PROGRAM MAIN
VAR

	fTotalCIP_Volume: REAL;
	fbWritePersistent: FB_WritePersistentData;
	bTesting		:	BOOL:=FALSE	;
	nI_1			: 	INT		;
	ftg_EStop_Fall	: 	F_TRIG	;
	rs_EStopFall	: 	RS	;
	bTestEstop		:	BOOL:=TRUE	;
	bTemp_Water_Overweight_check: BOOL;
	fbUPS: FB_S_UPS_CX51x0;

END_VAR

prg_RealClock();
prg_Piston();
prg_Safety();
prg_MessageManager();
prg_Messages();
prg_Call_OpMode();
prg_User();
act_ResetPumps();
(*
prg_TriBlender(
		fb_TriBlenderPump:= g_Pump.fbPump[E_Pump_List.TB0001],
		stTriblender:=stTriblender,
		arrComponents:=arrProductionComponents);
*)		
//act_SetAnalogSens_Test();//To be deleted, for testing purposes
act_Call_Sensors_Analog();//To be deleted, for testing purposes
act_Call_Sensors_Analog_1();//To be deleted, for testing purposes
act_Call_ScaleFactor();//To be deleted, for testing purposes
act_Call_ProcessCntrl();

act_Call_Pumps();
act_Sensors();
act_HeatExchenger();
//CIP <-> Siemens exchange
g_Anybus.fbSim(arToCip:=g_Anybus.arSimRaw, arFromCip:=gIO.Anybus_Outputs_Raw);
IF g_Anybus.bSimEnable THEN;
	g_Anybus.fbAnybus(bFieldbusOk:=TRUE, arRawIn:=g_Anybus.arSimRaw, arRawOut:=gIO.Anybus_Outputs_Raw);
ELSE;
	g_Anybus.fbAnybus(bFieldbusOk:=NOT gIO.Anybus_WcState, arRawIn:=gIO.Anybus_Inputs_Raw, arRawOut:=gIO.Anybus_Outputs_Raw);
END_IF
//Requests do not survive a PLC restart (Vadim, 02.11.2026)
IF NOT g_Anybus.bQueueCleared THEN;
	g_Data.fbCIP.m_PosDeleteAll_HMI();
	g_Anybus.bQueueCleared:=TRUE;
END_IF
IF g_Anybus.bBridgeEnable THEN;
	g_Anybus.fbBridge();
	g_Anybus.fbAnybus.stStatus:=g_Anybus.fbBridge.stStatus;
ELSE;
	g_Data.fbCIP.nLocalRecipe:=0;
END_IF
//One-time transfer of the old sets to the new recipes (Vadim 02.11.2026), the rest keeps the program defaults
IF g_Data.bRecipeTransfer THEN;
	g_Data.arr_CIP_Recipe[0]:=g_Data.arr_CIP_Param[E_CIP_Usage.eLocal];
	g_Data.arr_CIP_Recipe[1]:=g_Data.arr_CIP_Param[E_CIP_Usage.eTank_3];
	g_Data.arr_CIP_Recipe[2]:=g_Data.arr_CIP_Param[E_CIP_Usage.eLine_Color];
	g_Data.arr_CIP_Description[0]:='Local';
	g_Data.arr_CIP_Description[1]:='Tank - from Tank3 Color';
	g_Data.arr_CIP_Description[2]:='Pipe - from Line Color';
	g_Data.bRecipeTransfer:=FALSE;
END_IF
act_Call_CIP();

act_Call_For_HMI();

g_SFC.fbSFC_Temp1();

//Temtprary Overweght protection!!!!! DO NOT DELETE
IF fTotalCIP_Volume >=1500 AND FALSE THEN;
	//fbPis[E_Pis_Name.V1022].m_SetByRecipe(stPis:=stPis[E_Pis_Name.V1022], req:=E_Piston_Recipe_State.Release);
	//fbPis[E_Pis_Name.V1019].m_SetByRecipe(stPis:=stPis[E_Pis_Name.V1019], req:=E_Piston_Recipe_State.Release);
	//fbPis[E_Pis_Name.V1016].m_SetByRecipe(stPis:=stPis[E_Pis_Name.V1016], req:=E_Piston_Recipe_State.Release);
	//fbPis[E_Pis_Name.V1011].m_SetByRecipe(stPis:=stPis[E_Pis_Name.V1011], req:=E_Piston_Recipe_State.Release);
	bTemp_Water_Overweight_check:=FALSE;
	fbPrintErrMessageByID(sModuleDescription:='CIP',sActErrorID:='101x000x000');
ELSIF fTotalCIP_Volume < 1480 THEN;
	bTemp_Water_Overweight_check:=TRUE;
END_IF

IF arrTanksSens[E_Tank_Name.T91].get_stTankLevel_OverFlow() THEN;
	fbPis[E_Pis_Name.V1022].m_SetByRecipe(stPis:=stPis[E_Pis_Name.V1022], req:=E_Piston_Recipe_State.Release);
	//print error
	fbPrintErrMessageByID(sModuleDescription:='CIP',sActErrorID:='101x000x001');		
END_IF
IF arrTanksSens[E_Tank_Name.T92].get_stTankLevel_OverFlow() THEN;
	fbPis[E_Pis_Name.V1019].m_SetByRecipe(stPis:=stPis[E_Pis_Name.V1019], req:=E_Piston_Recipe_State.Release);
	//print error
	fbPrintErrMessageByID(sModuleDescription:='CIP',sActErrorID:='101x000x002');		
END_IF
IF arrTanksSens[E_Tank_Name.T93].get_stTankLevel_OverFlow() THEN;
	fbPis[E_Pis_Name.V1016].m_SetByRecipe(stPis:=stPis[E_Pis_Name.V1016], req:=E_Piston_Recipe_State.Release);
	//print error	
	fbPrintErrMessageByID(sModuleDescription:='CIP',sActErrorID:='101x000x003');	
END_IF
IF arrTanksSens[E_Tank_Name.T94].get_stTankLevel_OverFlow() THEN;
	fbPis[E_Pis_Name.V1011].m_SetByRecipe(stPis:=stPis[E_Pis_Name.V1011], req:=E_Piston_Recipe_State.Release);
	//print error
	fbPrintErrMessageByID(sModuleDescription:='CIP',sActErrorID:='101x000x004');		
END_IF
	


mElementList_SetName();

fbWritePersistent(
	NETID:= , 
	PORT:= 851, 
	START:= , 
	TMOUT:= T#3S, 
	MODE:= , 
	BUSY=> , 
	ERR=> , 
	ERRID=> );

fbUPS();

ACTION act_Call_CIP:
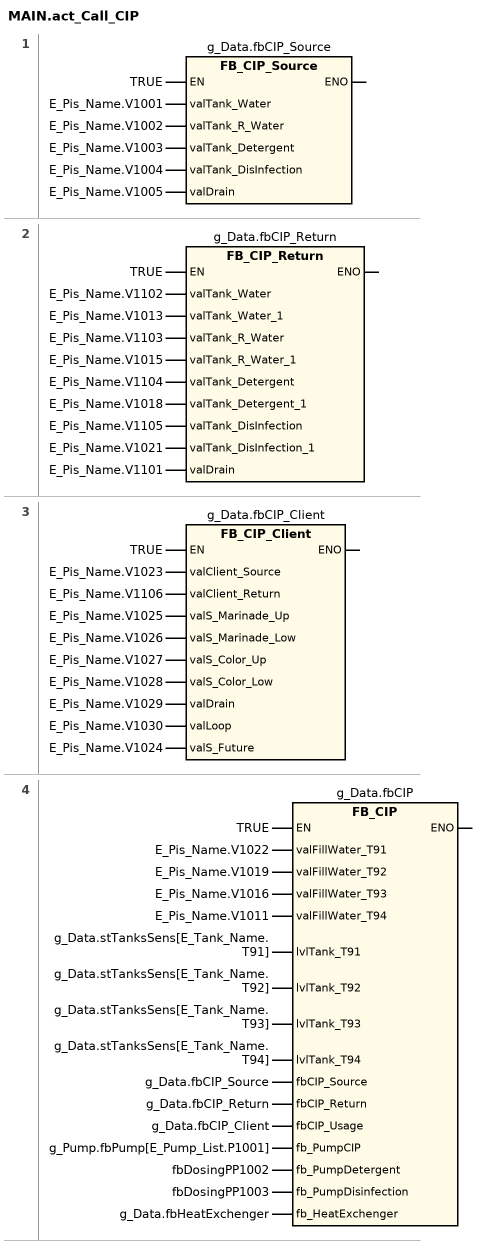
// NETWORK 1
g_Data.fbCIP_Source(
    valTank_Water := E_Pis_Name.V1001,
    valTank_R_Water := E_Pis_Name.V1002,
    valTank_Detergent := E_Pis_Name.V1003,
    valTank_DisInfection := E_Pis_Name.V1004,
    valDrain := E_Pis_Name.V1005); // FB_CIP_Source

// NETWORK 2
g_Data.fbCIP_Return(
    valTank_Water := E_Pis_Name.V1102,
    valTank_Water_1 := E_Pis_Name.V1013,
    valTank_R_Water := E_Pis_Name.V1103,
    valTank_R_Water_1 := E_Pis_Name.V1015,
    valTank_Detergent := E_Pis_Name.V1104,
    valTank_Detergent_1 := E_Pis_Name.V1018,
    valTank_DisInfection := E_Pis_Name.V1105,
    valTank_DisInfection_1 := E_Pis_Name.V1021,
    valDrain := E_Pis_Name.V1101); // FB_CIP_Return

// NETWORK 3
g_Data.fbCIP_Client(
    valClient_Source := E_Pis_Name.V1023,
    valClient_Return := E_Pis_Name.V1106,
    valS_Marinade_Up := E_Pis_Name.V1025,
    valS_Marinade_Low := E_Pis_Name.V1026,
    valS_Color_Up := E_Pis_Name.V1027,
    valS_Color_Low := E_Pis_Name.V1028,
    valDrain := E_Pis_Name.V1029,
    valLoop := E_Pis_Name.V1030,
    valS_Future := E_Pis_Name.V1024); // FB_CIP_Client

// NETWORK 4
g_Data.fbCIP(
    valFillWater_T91 := E_Pis_Name.V1022,
    valFillWater_T92 := E_Pis_Name.V1019,
    valFillWater_T93 := E_Pis_Name.V1016,
    valFillWater_T94 := E_Pis_Name.V1011,
    lvlTank_T91 := g_Data.stTanksSens[E_Tank_Name.T91],
    lvlTank_T92 := g_Data.stTanksSens[E_Tank_Name.T92],
    lvlTank_T93 := g_Data.stTanksSens[E_Tank_Name.T93],
    lvlTank_T94 := g_Data.stTanksSens[E_Tank_Name.T94],
    fbCIP_Source := g_Data.fbCIP_Source,
    fbCIP_Return := g_Data.fbCIP_Return,
    fbCIP_Usage := g_Data.fbCIP_Client,
    fb_PumpCIP := g_Pump.fbPump[E_Pump_List.P1001],
    fb_PumpDetergent := fbDosingPP1002,
    fb_PumpDisinfection := fbDosingPP1003,
    fb_HeatExchenger := g_Data.fbHeatExchenger); // FB_CIP
END_ACTION

ACTION act_Call_For_HMI:


g_HMI.stT91_Sens:=g_Data.stTanksSens[E_Tank_Name.T91];
g_HMI.stT92_Sens:=g_Data.stTanksSens[E_Tank_Name.T92];
g_HMI.stT93_Sens:=g_Data.stTanksSens[E_Tank_Name.T93];
g_HMI.stT94_Sens:=g_Data.stTanksSens[E_Tank_Name.T94];
END_ACTION

ACTION act_Call_ProcessCntrl:
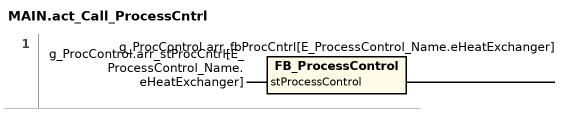
// NETWORK 1
g_ProcControl.arr_fbProcCntrl[E_ProcessControl_Name.eHeatExchanger](stProcessControl := g_ProcControl.arr_stProcCntrl[E_ProcessControl_Name.eHeatExchanger]); // FB_ProcessControl
END_ACTION

ACTION act_Call_Pumps:
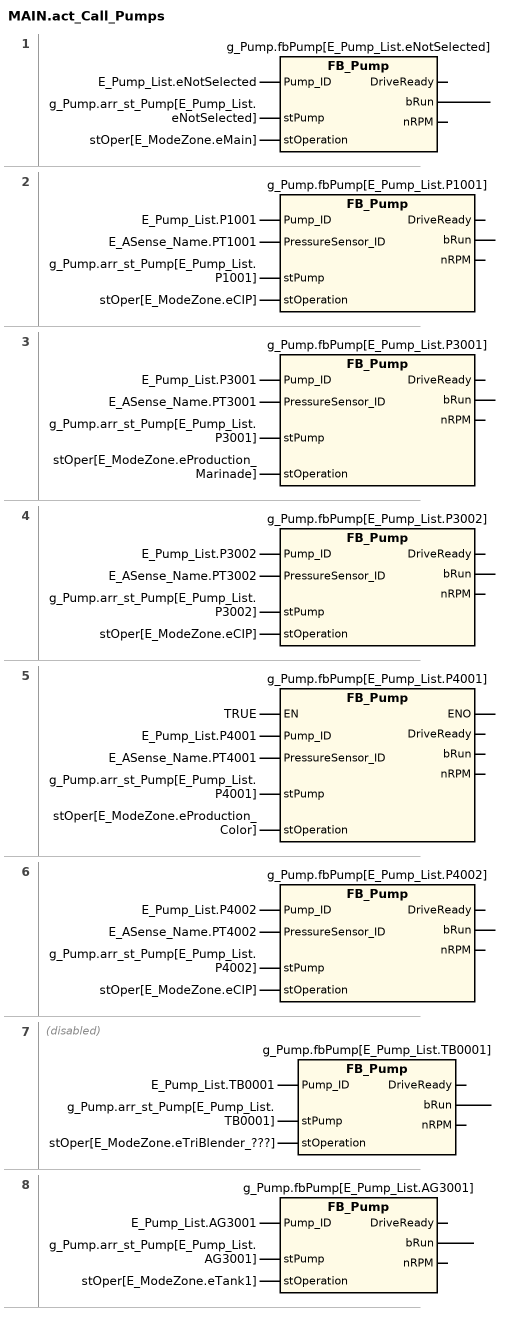
// NETWORK 1
g_Pump.fbPump[E_Pump_List.eNotSelected](
    Pump_ID := E_Pump_List.eNotSelected,
    stPump := g_Pump.arr_st_Pump[E_Pump_List.eNotSelected],
    stOperation := stOper[E_ModeZone.eMain]); // FB_Pump

// NETWORK 2
g_Pump.fbPump[E_Pump_List.P1001](
    Pump_ID := E_Pump_List.P1001,
    PressureSensor_ID := E_ASense_Name.PT1001,
    stPump := g_Pump.arr_st_Pump[E_Pump_List.P1001],
    stOperation := stOper[E_ModeZone.eCIP]); // FB_Pump

// NETWORK 3
g_Pump.fbPump[E_Pump_List.P3001](
    Pump_ID := E_Pump_List.P3001,
    PressureSensor_ID := E_ASense_Name.PT3001,
    stPump := g_Pump.arr_st_Pump[E_Pump_List.P3001],
    stOperation := stOper[E_ModeZone.eProduction_Marinade]); // FB_Pump

// NETWORK 4
g_Pump.fbPump[E_Pump_List.P3002](
    Pump_ID := E_Pump_List.P3002,
    PressureSensor_ID := E_ASense_Name.PT3002,
    stPump := g_Pump.arr_st_Pump[E_Pump_List.P3002],
    stOperation := stOper[E_ModeZone.eCIP]); // FB_Pump

// NETWORK 5
g_Pump.fbPump[E_Pump_List.P4001](
    Pump_ID := E_Pump_List.P4001,
    PressureSensor_ID := E_ASense_Name.PT4001,
    stPump := g_Pump.arr_st_Pump[E_Pump_List.P4001],
    stOperation := stOper[E_ModeZone.eProduction_Color]); // FB_Pump

// NETWORK 6
g_Pump.fbPump[E_Pump_List.P4002](
    Pump_ID := E_Pump_List.P4002,
    PressureSensor_ID := E_ASense_Name.PT4002,
    stPump := g_Pump.arr_st_Pump[E_Pump_List.P4002],
    stOperation := stOper[E_ModeZone.eCIP]); // FB_Pump

// NETWORK 7 (disabled)
// g_Pump.fbPump[E_Pump_List.TB0001](
//     Pump_ID := E_Pump_List.TB0001,
//     stPump := g_Pump.arr_st_Pump[E_Pump_List.TB0001],
//     stOperation := stOper[E_ModeZone.eTriBlender_???]); // FB_Pump

// NETWORK 8
g_Pump.fbPump[E_Pump_List.AG3001](
    Pump_ID := E_Pump_List.AG3001,
    stPump := g_Pump.arr_st_Pump[E_Pump_List.AG3001],
    stOperation := stOper[E_ModeZone.eTank1]); // FB_Pump

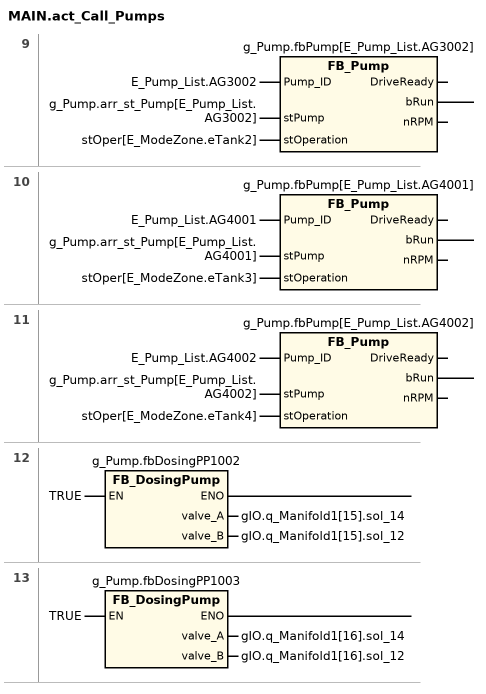
// NETWORK 9
g_Pump.fbPump[E_Pump_List.AG3002](
    Pump_ID := E_Pump_List.AG3002,
    stPump := g_Pump.arr_st_Pump[E_Pump_List.AG3002],
    stOperation := stOper[E_ModeZone.eTank2]); // FB_Pump

// NETWORK 10
g_Pump.fbPump[E_Pump_List.AG4001](
    Pump_ID := E_Pump_List.AG4001,
    stPump := g_Pump.arr_st_Pump[E_Pump_List.AG4001],
    stOperation := stOper[E_ModeZone.eTank3]); // FB_Pump

// NETWORK 11
g_Pump.fbPump[E_Pump_List.AG4002](
    Pump_ID := E_Pump_List.AG4002,
    stPump := g_Pump.arr_st_Pump[E_Pump_List.AG4002],
    stOperation := stOper[E_ModeZone.eTank4]); // FB_Pump

// NETWORK 12
g_Pump.fbDosingPP1002(valve_A => gIO.q_Manifold1[15].sol_14, valve_B => gIO.q_Manifold1[15].sol_12); // FB_DosingPump

// NETWORK 13
g_Pump.fbDosingPP1003(valve_A => gIO.q_Manifold1[16].sol_14, valve_B => gIO.q_Manifold1[16].sol_12); // FB_DosingPump
END_ACTION

ACTION act_Call_ScaleFactor:
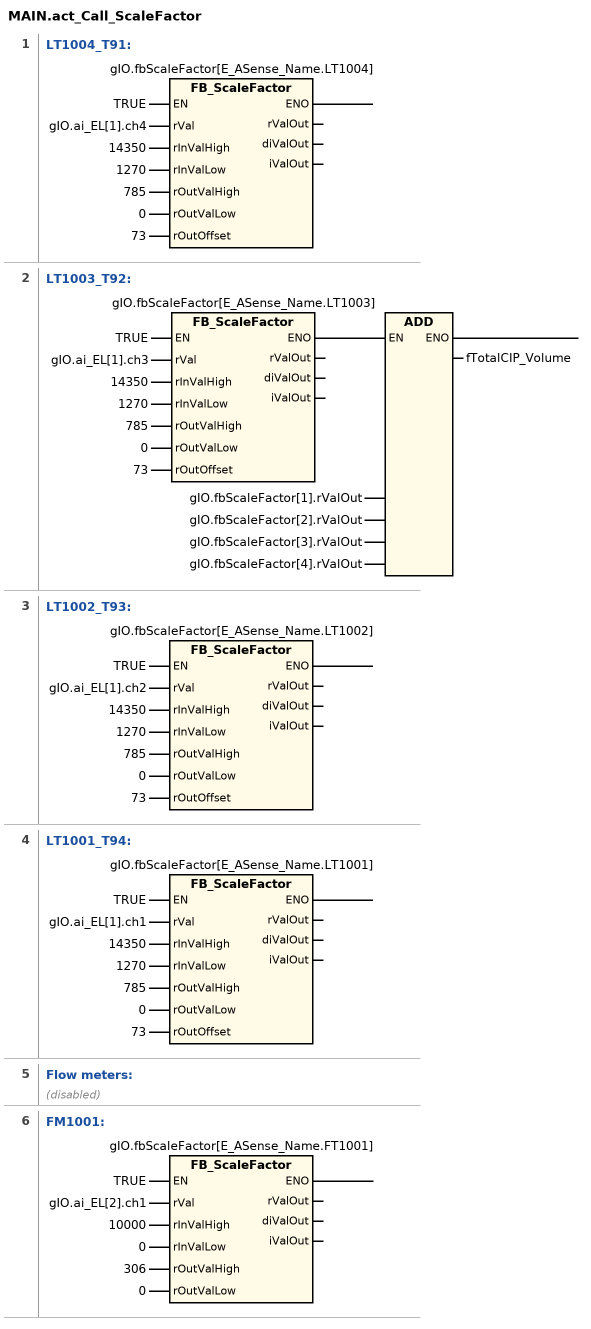
// NETWORK 1
LT1004_T91:
gIO.fbScaleFactor[E_ASense_Name.LT1004](
    rVal := gIO.ai_EL[1].ch4,
    rInValHigh := 14350,
    rInValLow := 1270,
    rOutValHigh := 785,
    rOutValLow := 0,
    rOutOffset := 73); // FB_ScaleFactor

// NETWORK 2
LT1003_T92:
gIO.fbScaleFactor[E_ASense_Name.LT1003](
    rVal := gIO.ai_EL[1].ch3,
    rInValHigh := 14350,
    rInValLow := 1270,
    rOutValHigh := 785,
    rOutValLow := 0,
    rOutOffset := 73); // FB_ScaleFactor
fTotalCIP_Volume := gIO.fbScaleFactor[1].rValOut + gIO.fbScaleFactor[2].rValOut + gIO.fbScaleFactor[3].rValOut + gIO.fbScaleFactor[4].rValOut;

// NETWORK 3
LT1002_T93:
gIO.fbScaleFactor[E_ASense_Name.LT1002](
    rVal := gIO.ai_EL[1].ch2,
    rInValHigh := 14350,
    rInValLow := 1270,
    rOutValHigh := 785,
    rOutValLow := 0,
    rOutOffset := 73); // FB_ScaleFactor

// NETWORK 4
LT1001_T94:
gIO.fbScaleFactor[E_ASense_Name.LT1001](
    rVal := gIO.ai_EL[1].ch1,
    rInValHigh := 14350,
    rInValLow := 1270,
    rOutValHigh := 785,
    rOutValLow := 0,
    rOutOffset := 73); // FB_ScaleFactor

// NETWORK 5 (disabled)
// label: Flow meters

// NETWORK 6
FM1001:
gIO.fbScaleFactor[E_ASense_Name.FT1001](
    rVal := gIO.ai_EL[2].ch1,
    rInValHigh := 10000,
    rInValLow := 0,
    rOutValHigh := 306,
    rOutValLow := 0); // FB_ScaleFactor

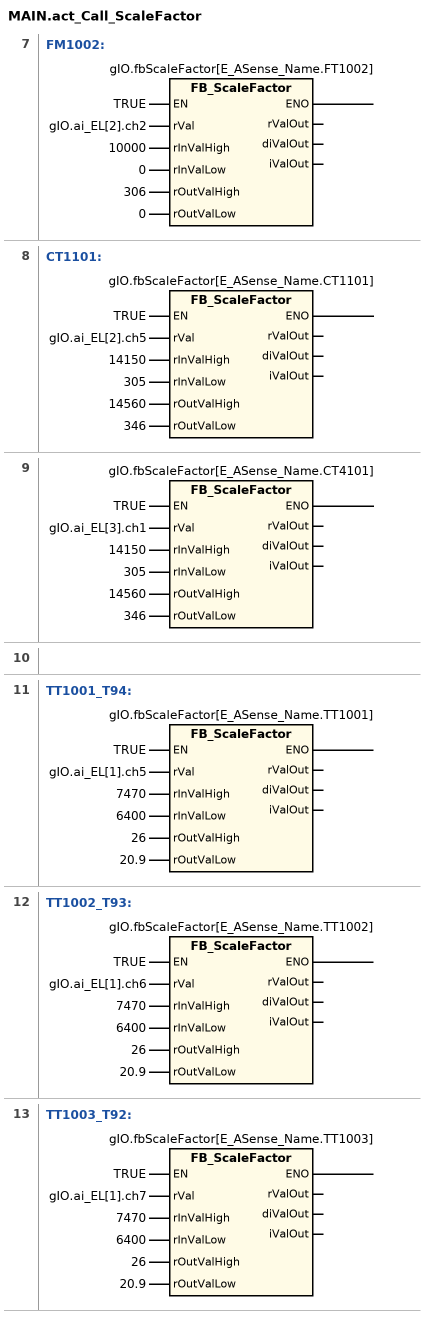
// NETWORK 7
FM1002:
gIO.fbScaleFactor[E_ASense_Name.FT1002](
    rVal := gIO.ai_EL[2].ch2,
    rInValHigh := 10000,
    rInValLow := 0,
    rOutValHigh := 306,
    rOutValLow := 0); // FB_ScaleFactor

// NETWORK 8
CT1101:
gIO.fbScaleFactor[E_ASense_Name.CT1101](
    rVal := gIO.ai_EL[2].ch5,
    rInValHigh := 14150,
    rInValLow := 305,
    rOutValHigh := 14560,
    rOutValLow := 346); // FB_ScaleFactor

// NETWORK 9
gIO.fbScaleFactor[E_ASense_Name.CT4101](
    rVal := gIO.ai_EL[3].ch1,
    rInValHigh := 14150,
    rInValLow := 305,
    rOutValHigh := 14560,
    rOutValLow := 346); // FB_ScaleFactor

// NETWORK 10

// NETWORK 11
TT1001_T94:
gIO.fbScaleFactor[E_ASense_Name.TT1001](
    rVal := gIO.ai_EL[1].ch5,
    rInValHigh := 7470,
    rInValLow := 6400,
    rOutValHigh := 26,
    rOutValLow := 20.9); // FB_ScaleFactor

// NETWORK 12
TT1002_T93:
gIO.fbScaleFactor[E_ASense_Name.TT1002](
    rVal := gIO.ai_EL[1].ch6,
    rInValHigh := 7470,
    rInValLow := 6400,
    rOutValHigh := 26,
    rOutValLow := 20.9); // FB_ScaleFactor

// NETWORK 13
TT1003_T92:
gIO.fbScaleFactor[E_ASense_Name.TT1003](
    rVal := gIO.ai_EL[1].ch7,
    rInValHigh := 7470,
    rInValLow := 6400,
    rOutValHigh := 26,
    rOutValLow := 20.9); // FB_ScaleFactor

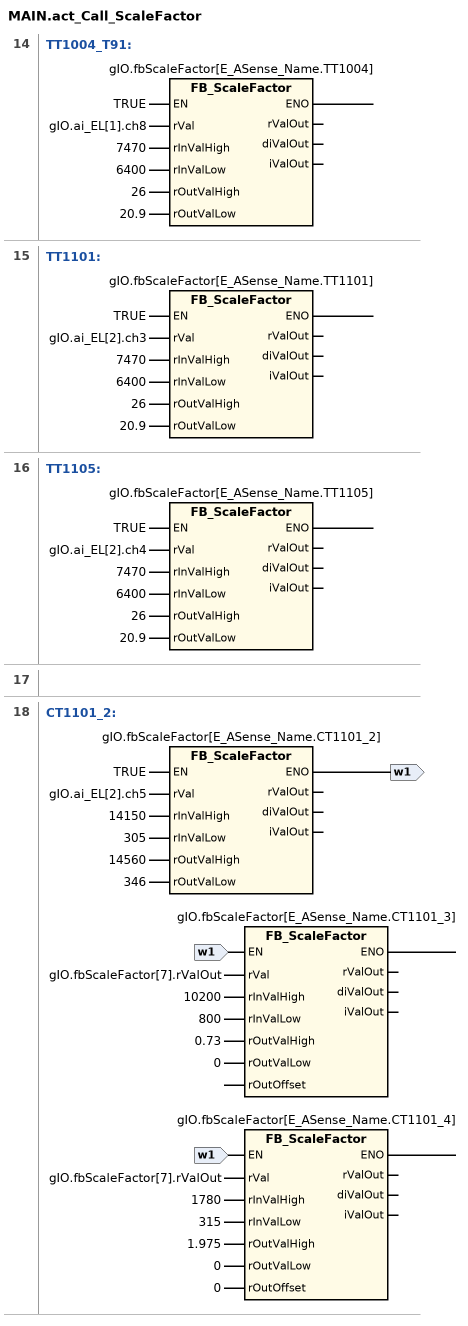
// NETWORK 14
TT1004_T91:
gIO.fbScaleFactor[E_ASense_Name.TT1004](
    rVal := gIO.ai_EL[1].ch8,
    rInValHigh := 7470,
    rInValLow := 6400,
    rOutValHigh := 26,
    rOutValLow := 20.9); // FB_ScaleFactor

// NETWORK 15
TT1101:
gIO.fbScaleFactor[E_ASense_Name.TT1101](
    rVal := gIO.ai_EL[2].ch3,
    rInValHigh := 7470,
    rInValLow := 6400,
    rOutValHigh := 26,
    rOutValLow := 20.9); // FB_ScaleFactor

// NETWORK 16
TT1105:
gIO.fbScaleFactor[E_ASense_Name.TT1105](
    rVal := gIO.ai_EL[2].ch4,
    rInValHigh := 7470,
    rInValLow := 6400,
    rOutValHigh := 26,
    rOutValLow := 20.9); // FB_ScaleFactor

// NETWORK 17

// NETWORK 18
CT1101_2:
gIO.fbScaleFactor[E_ASense_Name.CT1101_2](
    rVal := gIO.ai_EL[2].ch5,
    rInValHigh := 14150,
    rInValLow := 305,
    rOutValHigh := 14560,
    rOutValLow := 346); // FB_ScaleFactor
gIO.fbScaleFactor[E_ASense_Name.CT1101_3](
    rVal := gIO.fbScaleFactor[7].rValOut,
    rInValHigh := 10200,
    rInValLow := 800,
    rOutValHigh := 0.73,
    rOutValLow := 0); // FB_ScaleFactor
gIO.fbScaleFactor[E_ASense_Name.CT1101_4](
    rVal := gIO.fbScaleFactor[7].rValOut,
    rInValHigh := 1780,
    rInValLow := 315,
    rOutValHigh := 1.975,
    rOutValLow := 0,
    rOutOffset := 0); // FB_ScaleFactor

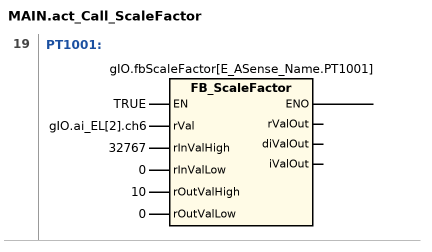
// NETWORK 19
PT1001:
gIO.fbScaleFactor[E_ASense_Name.PT1001](
    rVal := gIO.ai_EL[2].ch6,
    rInValHigh := 32767,
    rInValLow := 0,
    rOutValHigh := 10,
    rOutValLow := 0); // FB_ScaleFactor
END_ACTION

ACTION act_Call_Sensors_Analog:
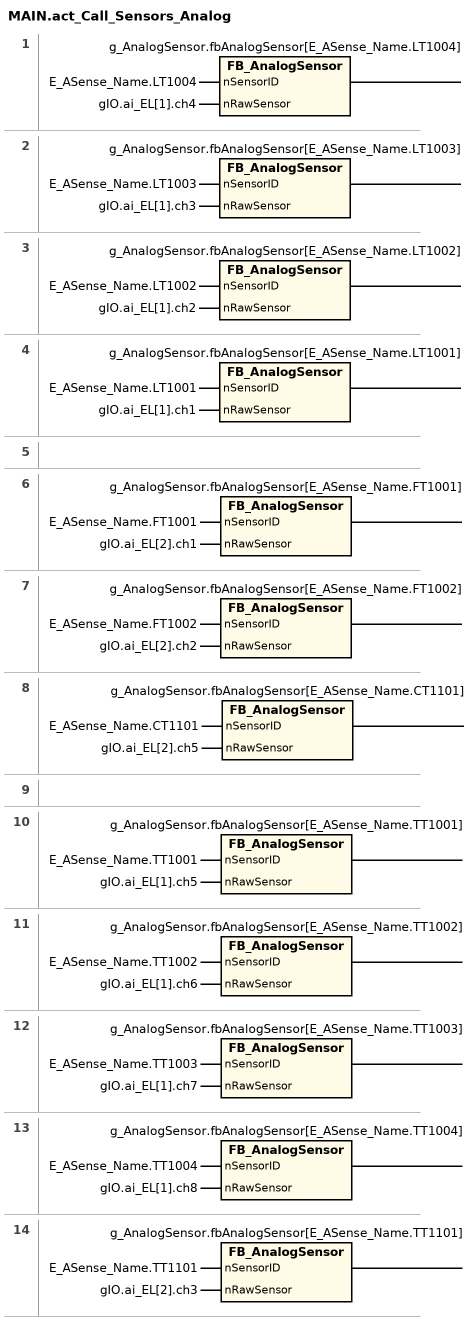
// NETWORK 1
g_AnalogSensor.fbAnalogSensor[E_ASense_Name.LT1004](nSensorID := E_ASense_Name.LT1004, nRawSensor := gIO.ai_EL[1].ch4); // FB_AnalogSensor

// NETWORK 2
g_AnalogSensor.fbAnalogSensor[E_ASense_Name.LT1003](nSensorID := E_ASense_Name.LT1003, nRawSensor := gIO.ai_EL[1].ch3); // FB_AnalogSensor

// NETWORK 3
g_AnalogSensor.fbAnalogSensor[E_ASense_Name.LT1002](nSensorID := E_ASense_Name.LT1002, nRawSensor := gIO.ai_EL[1].ch2); // FB_AnalogSensor

// NETWORK 4
g_AnalogSensor.fbAnalogSensor[E_ASense_Name.LT1001](nSensorID := E_ASense_Name.LT1001, nRawSensor := gIO.ai_EL[1].ch1); // FB_AnalogSensor

// NETWORK 5

// NETWORK 6
g_AnalogSensor.fbAnalogSensor[E_ASense_Name.FT1001](nSensorID := E_ASense_Name.FT1001, nRawSensor := gIO.ai_EL[2].ch1); // FB_AnalogSensor

// NETWORK 7
g_AnalogSensor.fbAnalogSensor[E_ASense_Name.FT1002](nSensorID := E_ASense_Name.FT1002, nRawSensor := gIO.ai_EL[2].ch2); // FB_AnalogSensor

// NETWORK 8
g_AnalogSensor.fbAnalogSensor[E_ASense_Name.CT1101](nSensorID := E_ASense_Name.CT1101, nRawSensor := gIO.ai_EL[2].ch5); // FB_AnalogSensor

// NETWORK 9

// NETWORK 10
g_AnalogSensor.fbAnalogSensor[E_ASense_Name.TT1001](nSensorID := E_ASense_Name.TT1001, nRawSensor := gIO.ai_EL[1].ch5); // FB_AnalogSensor

// NETWORK 11
g_AnalogSensor.fbAnalogSensor[E_ASense_Name.TT1002](nSensorID := E_ASense_Name.TT1002, nRawSensor := gIO.ai_EL[1].ch6); // FB_AnalogSensor

// NETWORK 12
g_AnalogSensor.fbAnalogSensor[E_ASense_Name.TT1003](nSensorID := E_ASense_Name.TT1003, nRawSensor := gIO.ai_EL[1].ch7); // FB_AnalogSensor

// NETWORK 13
g_AnalogSensor.fbAnalogSensor[E_ASense_Name.TT1004](nSensorID := E_ASense_Name.TT1004, nRawSensor := gIO.ai_EL[1].ch8); // FB_AnalogSensor

// NETWORK 14
g_AnalogSensor.fbAnalogSensor[E_ASense_Name.TT1101](nSensorID := E_ASense_Name.TT1101, nRawSensor := gIO.ai_EL[2].ch3); // FB_AnalogSensor

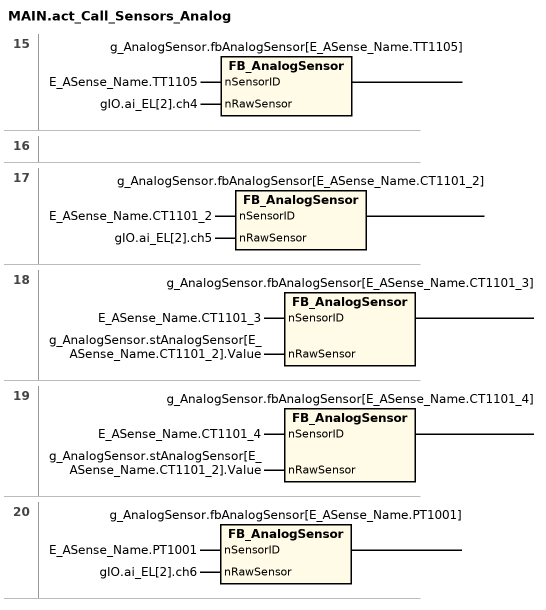
// NETWORK 15
g_AnalogSensor.fbAnalogSensor[E_ASense_Name.TT1105](nSensorID := E_ASense_Name.TT1105, nRawSensor := gIO.ai_EL[2].ch4); // FB_AnalogSensor

// NETWORK 16

// NETWORK 17
g_AnalogSensor.fbAnalogSensor[E_ASense_Name.CT1101_2](nSensorID := E_ASense_Name.CT1101_2, nRawSensor := gIO.ai_EL[2].ch5); // FB_AnalogSensor

// NETWORK 18
g_AnalogSensor.fbAnalogSensor[E_ASense_Name.CT1101_3](nSensorID := E_ASense_Name.CT1101_3, nRawSensor := g_AnalogSensor.stAnalogSensor[E_ASense_Name.CT1101_2].Value); // FB_AnalogSensor

// NETWORK 19
g_AnalogSensor.fbAnalogSensor[E_ASense_Name.CT1101_4](nSensorID := E_ASense_Name.CT1101_4, nRawSensor := g_AnalogSensor.stAnalogSensor[E_ASense_Name.CT1101_2].Value); // FB_AnalogSensor

// NETWORK 20
g_AnalogSensor.fbAnalogSensor[E_ASense_Name.PT1001](nSensorID := E_ASense_Name.PT1001, nRawSensor := gIO.ai_EL[2].ch6); // FB_AnalogSensor
END_ACTION

ACTION act_Call_Sensors_Analog_1:
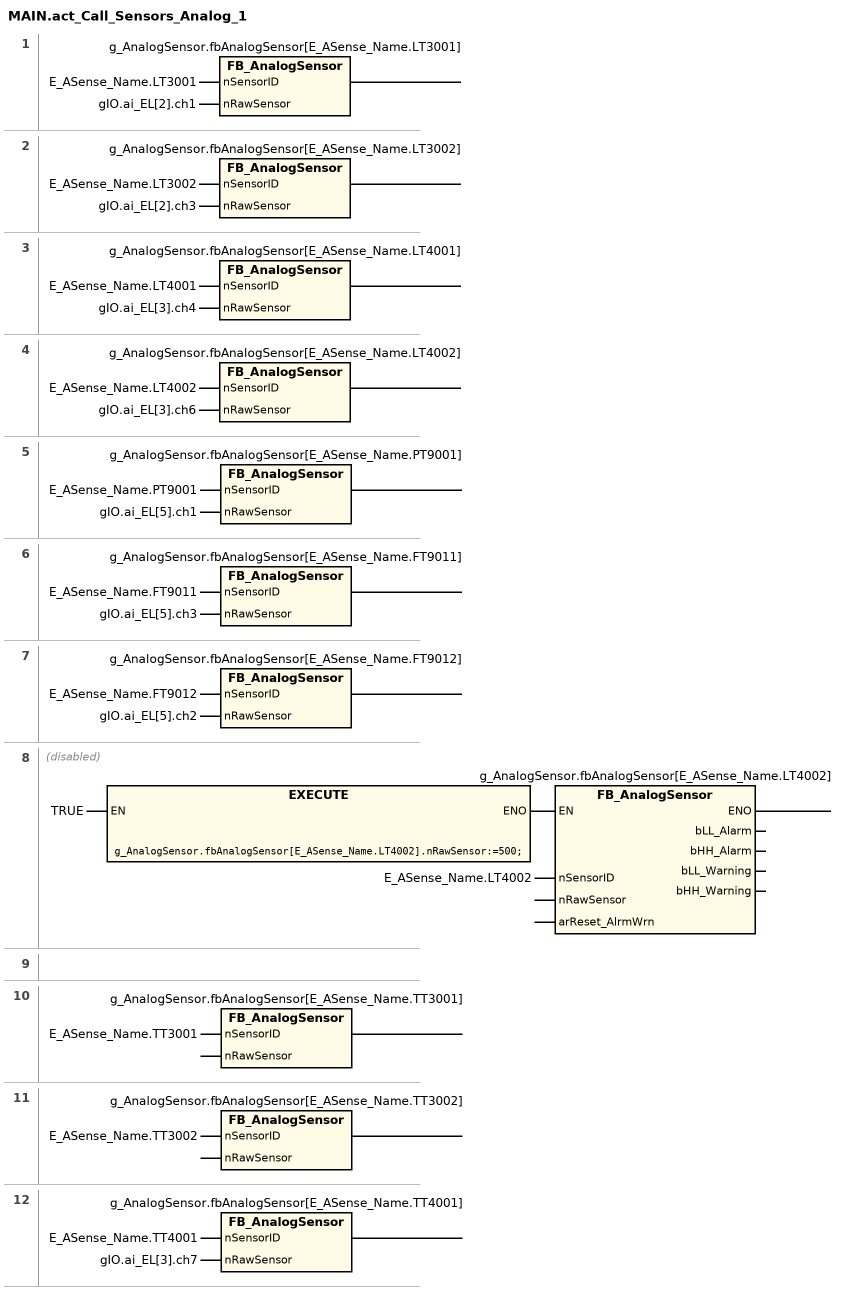
// NETWORK 1
g_AnalogSensor.fbAnalogSensor[E_ASense_Name.LT3001](nSensorID := E_ASense_Name.LT3001, nRawSensor := gIO.ai_EL[2].ch1); // FB_AnalogSensor

// NETWORK 2
g_AnalogSensor.fbAnalogSensor[E_ASense_Name.LT3002](nSensorID := E_ASense_Name.LT3002, nRawSensor := gIO.ai_EL[2].ch3); // FB_AnalogSensor

// NETWORK 3
g_AnalogSensor.fbAnalogSensor[E_ASense_Name.LT4001](nSensorID := E_ASense_Name.LT4001, nRawSensor := gIO.ai_EL[3].ch4); // FB_AnalogSensor

// NETWORK 4
g_AnalogSensor.fbAnalogSensor[E_ASense_Name.LT4002](nSensorID := E_ASense_Name.LT4002, nRawSensor := gIO.ai_EL[3].ch6); // FB_AnalogSensor

// NETWORK 5
g_AnalogSensor.fbAnalogSensor[E_ASense_Name.PT9001](nSensorID := E_ASense_Name.PT9001, nRawSensor := gIO.ai_EL[5].ch1); // FB_AnalogSensor

// NETWORK 6
g_AnalogSensor.fbAnalogSensor[E_ASense_Name.FT9011](nSensorID := E_ASense_Name.FT9011, nRawSensor := gIO.ai_EL[5].ch3); // FB_AnalogSensor

// NETWORK 7
g_AnalogSensor.fbAnalogSensor[E_ASense_Name.FT9012](nSensorID := E_ASense_Name.FT9012, nRawSensor := gIO.ai_EL[5].ch2); // FB_AnalogSensor

// NETWORK 8 (disabled)
// 
// 
// g_AnalogSensor.fbAnalogSensor[E_ASense_Name.LT4002].nRawSensor:=500;
// g_AnalogSensor.fbAnalogSensor[E_ASense_Name.LT4002](nSensorID := E_ASense_Name.LT4002); // FB_AnalogSensor

// NETWORK 9

// NETWORK 10
g_AnalogSensor.fbAnalogSensor[E_ASense_Name.TT3001](nSensorID := E_ASense_Name.TT3001); // FB_AnalogSensor

// NETWORK 11
g_AnalogSensor.fbAnalogSensor[E_ASense_Name.TT3002](nSensorID := E_ASense_Name.TT3002); // FB_AnalogSensor

// NETWORK 12
g_AnalogSensor.fbAnalogSensor[E_ASense_Name.TT4001](nSensorID := E_ASense_Name.TT4001, nRawSensor := gIO.ai_EL[3].ch7); // FB_AnalogSensor

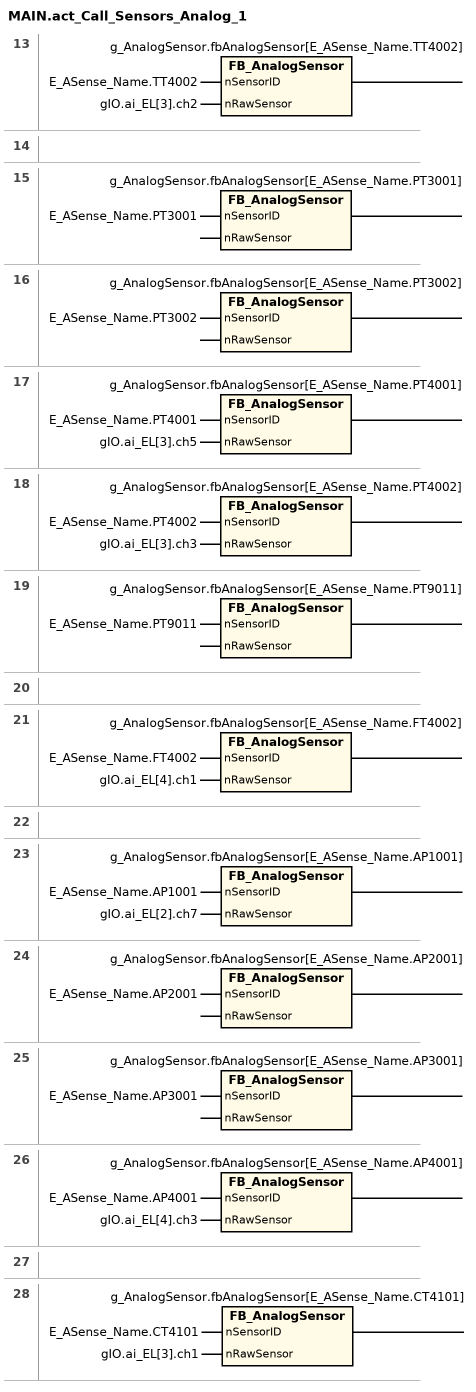
// NETWORK 13
g_AnalogSensor.fbAnalogSensor[E_ASense_Name.TT4002](nSensorID := E_ASense_Name.TT4002, nRawSensor := gIO.ai_EL[3].ch2); // FB_AnalogSensor

// NETWORK 14

// NETWORK 15
g_AnalogSensor.fbAnalogSensor[E_ASense_Name.PT3001](nSensorID := E_ASense_Name.PT3001); // FB_AnalogSensor

// NETWORK 16
g_AnalogSensor.fbAnalogSensor[E_ASense_Name.PT3002](nSensorID := E_ASense_Name.PT3002); // FB_AnalogSensor

// NETWORK 17
g_AnalogSensor.fbAnalogSensor[E_ASense_Name.PT4001](nSensorID := E_ASense_Name.PT4001, nRawSensor := gIO.ai_EL[3].ch5); // FB_AnalogSensor

// NETWORK 18
g_AnalogSensor.fbAnalogSensor[E_ASense_Name.PT4002](nSensorID := E_ASense_Name.PT4002, nRawSensor := gIO.ai_EL[3].ch3); // FB_AnalogSensor

// NETWORK 19
g_AnalogSensor.fbAnalogSensor[E_ASense_Name.PT9011](nSensorID := E_ASense_Name.PT9011); // FB_AnalogSensor

// NETWORK 20

// NETWORK 21
g_AnalogSensor.fbAnalogSensor[E_ASense_Name.FT4002](nSensorID := E_ASense_Name.FT4002, nRawSensor := gIO.ai_EL[4].ch1); // FB_AnalogSensor

// NETWORK 22

// NETWORK 23
g_AnalogSensor.fbAnalogSensor[E_ASense_Name.AP1001](nSensorID := E_ASense_Name.AP1001, nRawSensor := gIO.ai_EL[2].ch7); // FB_AnalogSensor

// NETWORK 24
g_AnalogSensor.fbAnalogSensor[E_ASense_Name.AP2001](nSensorID := E_ASense_Name.AP2001); // FB_AnalogSensor

// NETWORK 25
g_AnalogSensor.fbAnalogSensor[E_ASense_Name.AP3001](nSensorID := E_ASense_Name.AP3001); // FB_AnalogSensor

// NETWORK 26
g_AnalogSensor.fbAnalogSensor[E_ASense_Name.AP4001](nSensorID := E_ASense_Name.AP4001, nRawSensor := gIO.ai_EL[4].ch3); // FB_AnalogSensor

// NETWORK 27

// NETWORK 28
g_AnalogSensor.fbAnalogSensor[E_ASense_Name.CT4101](nSensorID := E_ASense_Name.CT4101, nRawSensor := gIO.ai_EL[3].ch1); // FB_AnalogSensor

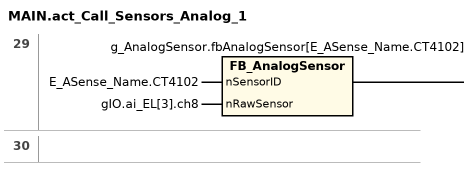
// NETWORK 29
g_AnalogSensor.fbAnalogSensor[E_ASense_Name.CT4102](nSensorID := E_ASense_Name.CT4102, nRawSensor := gIO.ai_EL[3].ch8); // FB_AnalogSensor

// NETWORK 30
END_ACTION

ACTION act_HeatExchenger:
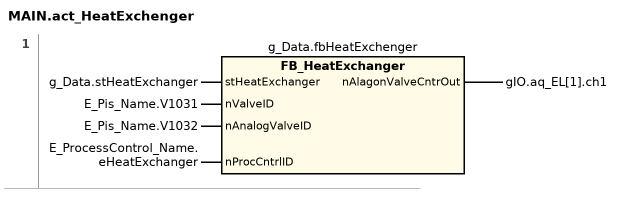
// NETWORK 1
g_Data.fbHeatExchenger(
    stHeatExchanger := g_Data.stHeatExchanger,
    nValveID := E_Pis_Name.V1031,
    nAnalogValveID := E_Pis_Name.V1032,
    nProcCntrlID := E_ProcessControl_Name.eHeatExchanger); // FB_HeatExchanger
gIO.aq_EL[1].ch1 := g_Data.fbHeatExchenger.nAlagonValveCntrOut;
END_ACTION

ACTION act_ResetPumps:
(*ftg_EStop_Fall(CLK:=prg_Safety.ftStateSafe.Q , Q=> );//EStop falling signal
rs_EStopFall(SET:=ftg_EStop_Fall.Q , RESET1:= , Q1=> );
IF rs_EStopFall.Q1 THEN
	FOR nI_1:=1 TO E_Pump_List.last BY 1 DO
		g_Pump.arr_st_Pump[nI_1].bRun_Auto:=FALSE;
	END_FOR
	rs_EStopFall.RESET1:=TRUE;
END_IF
rs_EStopFall.RESET1:=FALSE;*)
;
END_ACTION

ACTION act_Sensors:
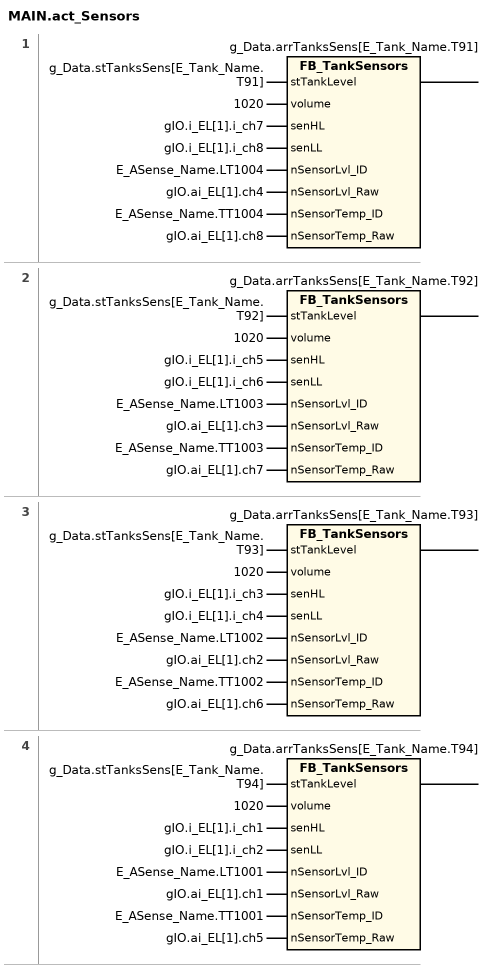
// NETWORK 1
g_Data.arrTanksSens[E_Tank_Name.T91](
    stTankLevel := g_Data.stTanksSens[E_Tank_Name.T91],
    volume := 1020,
    senHL := gIO.i_EL[1].i_ch7,
    senLL := gIO.i_EL[1].i_ch8,
    nSensorLvl_ID := E_ASense_Name.LT1004,
    nSensorLvl_Raw := gIO.ai_EL[1].ch4,
    nSensorTemp_ID := E_ASense_Name.TT1004,
    nSensorTemp_Raw := gIO.ai_EL[1].ch8); // FB_TankSensors

// NETWORK 2
g_Data.arrTanksSens[E_Tank_Name.T92](
    stTankLevel := g_Data.stTanksSens[E_Tank_Name.T92],
    volume := 1020,
    senHL := gIO.i_EL[1].i_ch5,
    senLL := gIO.i_EL[1].i_ch6,
    nSensorLvl_ID := E_ASense_Name.LT1003,
    nSensorLvl_Raw := gIO.ai_EL[1].ch3,
    nSensorTemp_ID := E_ASense_Name.TT1003,
    nSensorTemp_Raw := gIO.ai_EL[1].ch7); // FB_TankSensors

// NETWORK 3
g_Data.arrTanksSens[E_Tank_Name.T93](
    stTankLevel := g_Data.stTanksSens[E_Tank_Name.T93],
    volume := 1020,
    senHL := gIO.i_EL[1].i_ch3,
    senLL := gIO.i_EL[1].i_ch4,
    nSensorLvl_ID := E_ASense_Name.LT1002,
    nSensorLvl_Raw := gIO.ai_EL[1].ch2,
    nSensorTemp_ID := E_ASense_Name.TT1002,
    nSensorTemp_Raw := gIO.ai_EL[1].ch6); // FB_TankSensors

// NETWORK 4
g_Data.arrTanksSens[E_Tank_Name.T94](
    stTankLevel := g_Data.stTanksSens[E_Tank_Name.T94],
    volume := 1020,
    senHL := gIO.i_EL[1].i_ch1,
    senLL := gIO.i_EL[1].i_ch2,
    nSensorLvl_ID := E_ASense_Name.LT1001,
    nSensorLvl_Raw := gIO.ai_EL[1].ch1,
    nSensorTemp_ID := E_ASense_Name.TT1001,
    nSensorTemp_Raw := gIO.ai_EL[1].ch5); // FB_TankSensors
END_ACTION

ACTION act_SetAnalogSens_Test:
//set analog sensors setting only for the test. 
//Later this action should be deleted 
IF NOT bTesting THEN
	//Level
	g_AnalogSensor.stAnalogSensor[E_ASense_Name.LT1004].rawVal_Max:=14350;
	g_AnalogSensor.stAnalogSensor[E_ASense_Name.LT1004].rawVal_Min:=1270;
	g_AnalogSensor.stAnalogSensor[E_ASense_Name.LT1004].outVal_Max:=785;
	g_AnalogSensor.stAnalogSensor[E_ASense_Name.LT1004].outVal_Min:=0;
	g_AnalogSensor.stAnalogSensor[E_ASense_Name.LT1004].outOffset:=73;
	
	g_AnalogSensor.stAnalogSensor[E_ASense_Name.LT1003].rawVal_Max:=14350;
	g_AnalogSensor.stAnalogSensor[E_ASense_Name.LT1003].rawVal_Min:=1270;
	g_AnalogSensor.stAnalogSensor[E_ASense_Name.LT1003].outVal_Max:=785;
	g_AnalogSensor.stAnalogSensor[E_ASense_Name.LT1003].outVal_Min:=0;
	g_AnalogSensor.stAnalogSensor[E_ASense_Name.LT1003].outOffset:=73;
	
	g_AnalogSensor.stAnalogSensor[E_ASense_Name.LT1002].rawVal_Max:=14350;
	g_AnalogSensor.stAnalogSensor[E_ASense_Name.LT1002].rawVal_Min:=1270;
	g_AnalogSensor.stAnalogSensor[E_ASense_Name.LT1002].outVal_Max:=785;
	g_AnalogSensor.stAnalogSensor[E_ASense_Name.LT1002].outVal_Min:=0;
	g_AnalogSensor.stAnalogSensor[E_ASense_Name.LT1002].outOffset:=73;
	
	g_AnalogSensor.stAnalogSensor[E_ASense_Name.LT1001].rawVal_Max:=14350;
	g_AnalogSensor.stAnalogSensor[E_ASense_Name.LT1001].rawVal_Min:=1270;
	g_AnalogSensor.stAnalogSensor[E_ASense_Name.LT1001].outVal_Max:=785;
	g_AnalogSensor.stAnalogSensor[E_ASense_Name.LT1001].outVal_Min:=0;
	g_AnalogSensor.stAnalogSensor[E_ASense_Name.LT1001].outOffset:=73;
	
	//Flow
	g_AnalogSensor.stAnalogSensor[E_ASense_Name.FT1001].rawVal_Max:=10000;
	g_AnalogSensor.stAnalogSensor[E_ASense_Name.FT1001].rawVal_Min:=0;
	g_AnalogSensor.stAnalogSensor[E_ASense_Name.FT1001].outVal_Max:=306;
	g_AnalogSensor.stAnalogSensor[E_ASense_Name.FT1001].outVal_Min:=0;
	g_AnalogSensor.stAnalogSensor[E_ASense_Name.FT1001].outOffset:=0;
	
	g_AnalogSensor.stAnalogSensor[E_ASense_Name.FT1002].rawVal_Max:=10000;
	g_AnalogSensor.stAnalogSensor[E_ASense_Name.FT1002].rawVal_Min:=0;
	g_AnalogSensor.stAnalogSensor[E_ASense_Name.FT1002].outVal_Max:=306;
	g_AnalogSensor.stAnalogSensor[E_ASense_Name.FT1002].outVal_Min:=0;
	g_AnalogSensor.stAnalogSensor[E_ASense_Name.FT1002].outOffset:=0;
	
	////conductivity sensors
	g_AnalogSensor.stAnalogSensor[E_ASense_Name.CT1101].rawVal_Max:=14150;
	g_AnalogSensor.stAnalogSensor[E_ASense_Name.CT1101].rawVal_Min:=305;
	g_AnalogSensor.stAnalogSensor[E_ASense_Name.CT1101].outVal_Max:=14560;
	g_AnalogSensor.stAnalogSensor[E_ASense_Name.CT1101].outVal_Min:=346;
	g_AnalogSensor.stAnalogSensor[E_ASense_Name.CT1101].outOffset:=0;
	(*
	g_AnalogSensor.stAnalogSensor[E_ASense_Name.CT3101].rawVal_Max:=14150;
	g_AnalogSensor.stAnalogSensor[E_ASense_Name.CT3101].rawVal_Min:=305;
	g_AnalogSensor.stAnalogSensor[E_ASense_Name.CT3101].outVal_Max:=14560;
	g_AnalogSensor.stAnalogSensor[E_ASense_Name.CT3101].outVal_Min:=346;
	g_AnalogSensor.stAnalogSensor[E_ASense_Name.CT3101].outOffset:=0;
	*)
	//Temperature sensor
	g_AnalogSensor.stAnalogSensor[E_ASense_Name.TT1001].rawVal_Max:=7470;
	g_AnalogSensor.stAnalogSensor[E_ASense_Name.TT1001].rawVal_Min:=6400;
	g_AnalogSensor.stAnalogSensor[E_ASense_Name.TT1001].outVal_Max:=26;
	g_AnalogSensor.stAnalogSensor[E_ASense_Name.TT1001].outVal_Min:=20.9;
	g_AnalogSensor.stAnalogSensor[E_ASense_Name.TT1001].outOffset:=0;
	
	g_AnalogSensor.stAnalogSensor[E_ASense_Name.TT1002].rawVal_Max:=7470;
	g_AnalogSensor.stAnalogSensor[E_ASense_Name.TT1002].rawVal_Min:=6400;
	g_AnalogSensor.stAnalogSensor[E_ASense_Name.TT1002].outVal_Max:=26;
	g_AnalogSensor.stAnalogSensor[E_ASense_Name.TT1002].outVal_Min:=20.9;
	g_AnalogSensor.stAnalogSensor[E_ASense_Name.TT1002].outOffset:=0;
	
	g_AnalogSensor.stAnalogSensor[E_ASense_Name.TT1003].rawVal_Max:=7470;
	g_AnalogSensor.stAnalogSensor[E_ASense_Name.TT1003].rawVal_Min:=6400;
	g_AnalogSensor.stAnalogSensor[E_ASense_Name.TT1003].outVal_Max:=26;
	g_AnalogSensor.stAnalogSensor[E_ASense_Name.TT1003].outVal_Min:=20.9;
	g_AnalogSensor.stAnalogSensor[E_ASense_Name.TT1003].outOffset:=0;
	
	g_AnalogSensor.stAnalogSensor[E_ASense_Name.TT1004].rawVal_Max:=7470;
	g_AnalogSensor.stAnalogSensor[E_ASense_Name.TT1004].rawVal_Min:=6400;
	g_AnalogSensor.stAnalogSensor[E_ASense_Name.TT1004].outVal_Max:=26;
	g_AnalogSensor.stAnalogSensor[E_ASense_Name.TT1004].outVal_Min:=20.9;
	g_AnalogSensor.stAnalogSensor[E_ASense_Name.TT1004].outOffset:=0;
	
	g_AnalogSensor.stAnalogSensor[E_ASense_Name.TT1101].rawVal_Max:=7470;
	g_AnalogSensor.stAnalogSensor[E_ASense_Name.TT1101].rawVal_Min:=6400;
	g_AnalogSensor.stAnalogSensor[E_ASense_Name.TT1101].outVal_Max:=26;
	g_AnalogSensor.stAnalogSensor[E_ASense_Name.TT1101].outVal_Min:=20.9;
	g_AnalogSensor.stAnalogSensor[E_ASense_Name.TT1101].outOffset:=0;

	bTesting:=TRUE;
END_IF
END_ACTION

METHOD mElementList_SetName : BOOL
VAR_INPUT
END_VAR

VAR
	eASense_Name: E_ASense_Name;
	eProcCntrl: E_ProcessControl_Name;
END_VAR
FOR eASense_Name:=0 TO E_ASense_Name.last DO
	arAnalogSensorNameList[eASense_Name]:=TO_STRING(eASense_Name);
END_FOR

FOR eProcCntrl:=0 TO E_ProcessControl_Name.eProcCntrl_Last DO
	arr_ProcCntrl_NameList[eProcCntrl]:=TO_STRING(eProcCntrl);
	g_ProcControl.arr_stProcCntrl[eProcCntrl].idName:=TO_STRING(eProcCntrl);
END_FOR
END_METHOD

END_PROGRAM

(* stored: Version 1.1.0.1, ProductVersion 3.1.4026.21
   POU MAIN: Id {3441d04c-1b6a-45f8-92c9-effbc902d265}, SpecialFunc None
   Action act_Call_CIP: Id {23177538-beef-46ee-b17f-61590a7b02ee}
   Action act_Call_For_HMI: Id {95962895-82ce-49d5-9aef-33bffa18c9fd}
   Action act_Call_ProcessCntrl: Id {2101a6f8-5f32-44b3-875c-cd379d2d685c}
   Action act_Call_Pumps: Id {250d1796-6961-486b-9de7-1fb9e6e9ab7d}
   Action act_Call_ScaleFactor: Id {774d29d4-9ded-47dd-863a-e1e521c0ad31}
   Action act_Call_Sensors_Analog: Id {7ffdbc56-05dc-45ee-9e2a-e9c205335a24}
   Action act_Call_Sensors_Analog_1: Id {c3b256f4-619a-4513-b623-368be1d897cc}
   Action act_HeatExchenger: Id {bf3394df-98fc-4323-89aa-f243bd329b49}
   Action act_ResetPumps: Id {d6d5f25f-7520-4a69-86f1-bc96d10af8f9}
   Action act_Sensors: Id {8d3d0c01-4d42-45d2-a1c2-ec56cd1d1464}
   Action act_SetAnalogSens_Test: Id {455abcb0-c90c-4f45-9ea9-f7b3ab53cef4}
   Method mElementList_SetName: Id {fee97784-09c9-4c65-955f-9f389d44d720} *)
